// TwinCAT 3 PLC project Weegschaal
// ProgramVersion: 3.1.4024.0
// libraries:
//   Tc2_SerialCom, * (Beckhoff Automation GmbH)
//   Tc2_Standard, * (Beckhoff Automation GmbH)
//   Tc2_System, * (Beckhoff Automation GmbH)
//   Tc3_Module, * (Beckhoff Automation GmbH)
// project tree:
//   DUTs/ FB_ParseWeight.TcPOU
//   GVLs/ GVL.TcGVL
//   / PlcTask.TcTTO
//   POUs/ MAIN.TcPOU
// real-time tasks:
//   TASK PlcTask: cycle T#10ms, priority 20, ADS port 350
// I/O:
//   DEVICE Device 1 (EtherCAT), AmsNetId 5.59.220.46.2.1
//     Term 1 (EK1200) [EK1200-5000 EtherCAT Power supply (2A E-Bus)]
//       Term 2 (EL1008) [EL1008 8Ch. Dig. Input 24V, 3ms]
//       Term 3 (EL2008) [EL2008 8Ch. Dig. Output 24V, 0.5A]
//       Term 4 (EL3062) [EL3062 2Ch. Ana. Input 0-10V]
//       Term 5 (EL4002) [EL4002 2Ch. Ana. Output 0-10V, 12bit]
//       Term 6 (EK1110) [EK1110 EtherCAT extension]
//   DEVICE Device 3 (EtherCAT), AmsNetId 5.59.220.46.4.1
//     Term 7 (EK1100) [EK1100 EtherCAT Coupler (2A E-Bus)]
//       Term 8 (EL6851) [EL6851 DMX Master]
//       Term 9 (EL6002) [EL6002 Interface 2Ch. (RS232)]
//       Term 4 (EL9011) [EL9011 End Terminal]
//   DEVICE Device 2 (NOV-DP-RAM)
// variable links:
//   Weegschaal/Weegschaal Instance <-> Device 3 (EtherCAT)/Term 7 (EK1100)/Term 9 (EL6002)
//     PlcTask Inputs/GVL.stEL6002_In/D <-> COM TxPDO-Map Inputs Channel 2/Data In 0
//     PlcTask Inputs/GVL.stEL6002_In/D @bit {8..168 step 8} <-> COM TxPDO-Map Inputs Channel 2/Data In {1..21}  (21 links)
//     PlcTask Inputs/GVL.stEL6002_In/Status <-> COM TxPDO-Map Inputs Channel 2/Status
//     PlcTask Outputs/GVL.stEL6002_Out/Ctrl <-> COM RxPDO-Map Outputs Channel 2/Ctrl
//     PlcTask Outputs/GVL.stEL6002_Out/D <-> COM RxPDO-Map Outputs Channel 2/Data Out 0
//     PlcTask Outputs/GVL.stEL6002_Out/D @bit {8..168 step 8} <-> COM RxPDO-Map Outputs Channel 2/Data Out {1..21}  (21 links)

CONFIGURATION Weegschaal
    RESOURCE PLC ON TwinCAT3
        TASK PlcTask(INTERVAL := T#10ms, PRIORITY := 20);
        PROGRAM MAIN WITH PlcTask : MAIN;
    END_RESOURCE
END_CONFIGURATION

// ---- GVLs/GVL.TcGVL
VAR_GLOBAL
    // Correct Data Types for EL60xx Terminals in 22-byte mode
    stEL6002_In  AT %I* : EL6inData22B;  // "i" is lowercase in the official type name
    stEL6002_Out AT %Q* : EL6outData22B; // "o" is lowercase in the official type name
    
    RxBuffer : ComBuffer;
    TxBuffer : ComBuffer;
END_VAR

// ---- POUs/MAIN.TcPOU
PROGRAM MAIN
VAR
    // Serial communication blocks
    fbSerialLineControl : SerialLineControl;
    fbReceiveString     : ReceiveString;
    fbParseWeight       : FB_ParseWeight; 
    
    // Communication variables
    sRawData            : STRING(255);
    bStringReceived     : BOOL;
    bRxBusy             : BOOL;
    bRxError            : BOOL;
    nRxErrorID          : UDINT;
    
    // Parsing results
    fCurrentWeight      : LREAL;
    sUnit               : STRING(3);
    bDataValid          : BOOL;
    
    // Stability results
    bStableReading      : BOOL;
    fLastStableWeight   : LREAL;
END_VAR

// ==========================================================
// 1. BACKGROUND COMMUNICATION (Run this every cycle)
// ==========================================================
fbSerialLineControl(
    Mode        := SERIALLINEMODE_EL6_22B,
    pComIn      := ADR(stEL6002_In),
    pComOut     := ADR(stEL6002_Out),
    SizeComIn   := SIZEOF(stEL6002_In),
    TxBuffer    := TxBuffer,
    RxBuffer    := RxBuffer
);

// ==========================================================
// 2. RECEIVE CONTINUOUS STREAM DATA
// ==========================================================
fbReceiveString(
    Prefix          := '',
    Suffix          := '$R$N',
    Timeout         := T#1S,
    ReceivedString  := sRawData,
    RxBuffer        := RxBuffer,
    StringReceived  => bStringReceived,
    Busy            => bRxBusy
);

// ==========================================================
// 3. PARSE AND CHECK STABILITY (Alleen bij nieuwe data)
// ==========================================================
IF bStringReceived THEN
    fbParseWeight(
        sRawData            := sRawData,
        fStabilityThreshold := 0.001,
        fCurrentWeight      => fCurrentWeight,
        sUnit               => sUnit,
        bStableReading      => bStableReading,
        fLastStableWeight   => fLastStableWeight,
        bDataValid          => bDataValid
    );
END_IF

END_PROGRAM

// ---- DUTs/FB_ParseWeight.TcPOU
FUNCTION_BLOCK FB_ParseWeight
VAR_INPUT
    sRawData            : STRING(255);
    fStabilityThreshold : LREAL := 0.001;
END_VAR
VAR_OUTPUT
    fCurrentWeight      : LREAL;
    sUnit               : STRING(3);
    bStableReading      : BOOL;
    fLastStableWeight   : LREAL;
    bDataValid          : BOOL;
END_VAR
VAR
    sWeightTrimmed      : STRING(255);
    sSign               : STRING(1);
    aReadings           : ARRAY[1..5] OF LREAL;
    i                   : INT;
    fMaxReading         : LREAL;
    fMinReading         : LREAL;
END_VAR

// Initialisatie
bDataValid := FALSE;

// Controleer of er voldoende data is
IF LEN(sRawData) >= 10 THEN
    
    // Extract Sign (Position 1)
    sSign := MID(sRawData, 1, 1);
    
    // Extract Weight Value (Positions 3 to 9)
    sWeightTrimmed := MID(sRawData, 7, 3);
    
    // Remove blank spaces in the string
    sWeightTrimmed := REPLACE(sWeightTrimmed, '', 1, FIND(sWeightTrimmed, ' '));
    
    // Convert to floating point
    fCurrentWeight := TO_LREAL(sWeightTrimmed);
    
    // Apply negative sign if necessary
    IF sSign = '-' THEN
        fCurrentWeight := fCurrentWeight * -1.0;
    END_IF
    
    // Extract Unit (Positions 11 to 12)
    sUnit := MID(sRawData, 2, 11);
    
    // ==========================================================
    // STABILITY CHECK
    // ==========================================================
    // Shift old readings left
    FOR i := 1 TO 4 DO
        aReadings[i] := aReadings[i+1];
    END_FOR
    aReadings[5] := fCurrentWeight; // Append new reading
    
    // Calculate Min and Max in the buffer
    fMinReading := aReadings[1];
    fMaxReading := aReadings[1];
    FOR i := 2 TO 5 DO
        IF aReadings[i] < fMinReading THEN fMinReading := aReadings[i]; END_IF;
        IF aReadings[i] > fMaxReading THEN fMaxReading := aReadings[i]; END_IF;
    END_FOR
    
    // Evaluate threshold
    IF (fMaxReading - fMinReading) <= fStabilityThreshold THEN
        bStableReading := TRUE;
        fLastStableWeight := fCurrentWeight;
    ELSE
        bStableReading := FALSE;
    END_IF
    
    bDataValid := TRUE;
    
END_IF

END_FUNCTION_BLOCK
